(* IEC 61131-3 sources: JingjiangArm/moonboxpro_arm_8.4/Application/Application/任务列表/LogTask/文件存储/数据存储&日志操作, 8 files *)

(* ---- ENUMS_TIMEFORMAT.st ---- *)
(*@CES
Name=ENUMS_TIMEFORMAT
Type=Gvl
TypeGuid=2db5746d-d284-4425-9f7f-2663a34b0ebc
Guid=3fd86c5d-f4c2-4e63-8cc9-6ae2cca08ccd
HasDeclaration=True
HasImplementation=False
*)
{DECLARATION}
//{attribute 'qualified_only'}
//{attribute 'strict'}
TYPE ENUMS_TIMEFORMAT : (
	TIMEFORMAT_NO_HYPHEN		, (* yyyymmddHHMMSS *)
	TIMEFORMAT_HYPHEN_COLON		, (* yyyy-mm-dd HH:MM:SS *)
	TIMEFORMAT_HYPHEN_DOT		, (* yyyy.mm.dd.HHMMSS *)
	TIMEFORMAT_MMDD				, (* mmdd *)
	TIMEFORMAT_MMDDHH			  (* mmddHH *)
);
END_TYPE
{IMPLEMENTATION}

(* ---- StAxisWatchDetails.st ---- *)
(*@CES
Name=StAxisWatchDetails
Type=Gvl
TypeGuid=2db5746d-d284-4425-9f7f-2663a34b0ebc
Guid=06521707-3ba7-4049-9244-d2161cd79c22
HasDeclaration=True
HasImplementation=False
*)
{DECLARATION}
{attribute 'pack_mode' := '1'}
TYPE StAxisWatchDetails :
STRUCT
// 	iStationId						: INT;(*主控站ID*)
// 	rGirth 							:REAL ; (*周长*)
// 	iRtn_Station					: INT;//返回值
// 	iRunMode_Station				: INT;//运动模式-3电子齿轮4龙门
// 	rPos_Prf						: REAL;//规划位置
// 	rPos_Enc						: REAL;//编码器位置
// 	rVel_Enc						: REAL;//编码器速度
// 	rTorque							: REAL;//扭矩输出
// 	rGantry_Err						: REAL;//龙门错误吗
//  	rTemperaTure					: REAL;//电机温度
// 	dwErr_Driver					: DWORD;//驱动器报警状态
// 	wSts_Driver						: WORD;//驱动器状态
// 	wSts_NetPort					: WORD;//端口状态
// 	wSts_NetRun						: WORD;//端口运行状态
//  	iErr_NetPort_a					: INT;//A误码率
//  	iErr_NetPort_b					: INT;//B误码率
// 	dwMotion_Sts					: DWORD;//运型状态
// 	uiVirtual_Cnt					: UINT;//虚拟码盘基数
// 	wVirtual_Sts					: WORD;//虚拟马盘状态
// 	uiBrake_Cnt						: UINT;//制动次数
// 	rCurrent_Driver					: REAL;//电流
// 	rVdc							: REAL;//母线电压
// 	uiStationType					: UINT;//站类型
// 	uiDrvParam_Imax					: UINT;(* 驱动参数|最大电流 *)
// 	uiDrvParam_Nrs					: UINT;(* 驱动参数|额定转速 *)
// 	uiDrvParam_Nos					: UINT;(* 驱动参数|过速转速 *)
// 	iDrvParam_PosOfst				: INT;(* 驱动参数|位置偏移 *)

	rGirth: REAL; (* 轴周长 *)
	lrPT_Pos: LREAL; (* 轴PT规划P *)
	diPT_Time: DINT; (* 轴PT规划T *)
	byPT_Type: BYTE; (* 轴PT段选择|2.PT_SEGMENT_NORMAL;1.PT_SEGMENT_EVEN;0.others *)
	rtnSts: INT; (* 返回状态 *)
	bySpace: BYTE; (* fifo空间 *)
	pfr: DWORD; (* 规划位置 *)
	enc_Lo16: INT; (* StPTSts.enc的低16位_跟随误差的低16位 *)
	driverSts: INT; (* 驱动器状态 *)
	driverErr: INT; (* 驱动器错误 *)
	netPortErr_a: INT; (* A口误码率 *)
	netPortErr_b: INT; (* B口误码率 *)
	motionSts: DWORD; (* 运动器状态 *)
	modal: WORD; (* 模态 *)
	brakeCnt: WORD; (* 制动电阻次数 *)
	driverCurrent: WORD; (* 驱动器电流 *)
	rVel_Axis: REAL; (* 轴速度 *)
	rAI_Axis_Coating: REAL; (* 当前值-中位值 *)
	enc_Hi16: WORD; (* StPTSts.enc的高16位_网络锁存时间的低16位 *)(* 新增14个字节|@2020.10.13.171810_ *)
	temperature: INT; (* 电机温度 *)
	vel: INT; (* 规划速度 *)
	netPortSts: INT; (* 网络端口连接状态 *)
	netRunSts: INT; (* 网络运行状态 *)
	virtualCnt: WORD; (* 虚拟码盘计数 *)
	virtualSts: WORD; (* 虚拟码盘状态 *)
	(*2022.5.25.131916 增加了锁存编码器值的保存*)
	dwCurAxisEnc_Lock: DWORD;(*当前轴锁存编码器值*)
	dwCurAxisSystime_Lock					: DWORD;(*当前轴锁存系统时间*)
(*2022.6.24.151851  取消使用*)
(*
	dwLastLinkageAxisEnc_Lock				: DWORD;(*上个联动轴锁存编码器值*)
	dwLastLinkageAxisSystime_Lock			: DWORD;(*上个联动轴锁存系统时间*)
*)
	(*2022.6.24.151255*)
	iai1_New16D:			INT;(*模拟量输入1*)
	iai2_New16D:			INT;(*温控输入*)
	rDc_Voltage:REAL;(*母线电压值*)
	idriverErr_H: INT; (* 驱动器错误 |高16bit*)

	(*新增加的单联动切换功能，在出现问题的时候为了方便查找问题,增加了文件保存内容*)
	(*电机使能模式|0: 不使能 1: 使能 3: 使能后轴可以手动转动 4: 取消模式3状态
	3、4以为的值都不允许set
	实际应用下会3、4状态下切换*)
	wEnableMode_Motor						: WORD;
	byEnableModeSwitchDne					: BYTE;(*使能模式切换成功了|.0 =3 成功了
																		.1 =4 成功了*)
	xMoveEnable_Motor						: BOOL;(*电机运动使能|用于控制驱动器是否进行电机控制|与单联动比较切换电机是否运动*)

	byAxisMotionSts:BYTE;(*轴运动状态标志|0:同步运动状态.
										  |1:同步运动时停止运动状态.
										  |2:停止运动状态
										  |3:停止运动时加速到单运行速度状态.
										  |4:单运行时减速到停止状态.
										  |5:停止运动时或者使用单运行速度运行时加速到同步运动状态.
										  |6:非同步运动时急停到0状态.
										  |7:非同步运动时空转停机到0状态.*)
(*2022.10.22.162829保存加热相关数据*)
	rPIDValue:REAL;(*pid计算调整量*)
	rPV_Unit:REAL;(*当前温度*)
	rSV_Unit:REAL;(*设定温度*)
	rValue_P:REAL;
	rValue_I:REAL;
	rValue_D:REAL;
	iNumCount:INT;

(*end_2022.10.22.163310*)

END_STRUCT
END_TYPE

{IMPLEMENTATION}

(* ---- StRecord_A.st ---- *)
(*@CES
Name=StRecord_A
Type=Gvl
TypeGuid=2db5746d-d284-4425-9f7f-2663a34b0ebc
Guid=136b24a0-c4f1-416e-bf48-48716262a31a
HasDeclaration=True
HasImplementation=False
*)
{DECLARATION}
{attribute 'pack_mode' := '1'}
TYPE StRecord_A :
STRUCT
	dwCurYMD: DWORD;
	dwCurHMSU: DWORD;
	byAxisId: BYTE; (* 轴id *)
	byGrpId: BYTE; (* 系id *)
	uiNum: UINT; (* 减速比分子 *)
	uiDen: UINT; (* 减速比分母 *)
	udiVel: UDINT; (* 主机速度|单位:0.01m/min *)
	udiGirth: UDINT; (* 版周长|单位:0.001mm *)
	iGateSa: INT; (* 波门地址1 *)
	iGateSaEx: INT; (* 波门地址2 *)
	byMarkTypeId: BYTE; (* 标记形式 *)
	byMarkArrangeId: BYTE; (* 标记排列 *)
	wSwitchRef: WORD; (* 开关状态 *)
	wStatusRef: WORD; (* 手/自动状态 *)
	wExtendedProf: WORD;
			(* 描述位|
				bit0=1表示合压中,
				bit1=1标识等料长,
				bit2=1标识裁切让料头

				bit8=1表示第一组波门T1极性
				bit9=1表示第一组波门T2极性
				bit10=1表示第二组波门T1极性
				bit11=1表示第二组波门T2极性
*)
	byStsV: BYTE; (* 纵向误差状态 *)
	byStsH: BYTE; (* 横向误差状态 *)
	aiKpid_setup_v: ARRAY [1..3] OF INT; (*界面设置的纵向pid*)
	aiKpid_setup_h: ARRAY [1..3] OF INT; (*界面设置的横向pid*)
	aiKpid_used_v: ARRAY [1..3] OF INT; (*使用中的纵向pid*)
	aiAdjVal_vh: ARRAY [1..2] OF INT; (*纵横向版修正量*)
	lrFilmLengthFromPrevUnit: LREAL; (* 预套准料长总值 *)
	byCouplingMask: BYTE; (* 耦合开关 *)
	iErrDataRelay_Index_V: INT; (* 取的误差间隔幅数 *)
	iErrDataRelay_V: INT; (* 传来的误差 *)
	aiErrorVal_vh: ARRAY [1..2] OF INT; (*纵横向误差*)
	aiAdjValCalcByPid_vh: ARRAY [1..2] OF INT; (*计算的调整量*)

	alrCurCycleAdjustVal_Auto_vh: ARRAY [1..2] OF LREAL; (* 自动调整*)
	alrCurCycleAdjustVal_Rapid_vh: ARRAY [1..2] OF LREAL; (* 快速对版调整*)
	alrCurCycleAdjustVal_ManuCoarse_vh: ARRAY [1..2] OF LREAL; (* 手动粗调*)
	alrCurCycleAdjustVal_ManuFine_vh: ARRAY [1..2] OF LREAL; (* 手动细调*)
	alrCurCycleAdjustVal_Coupling_vh: ARRAY [1..2] OF LREAL; (* 耦合量*)
	alrCurcycleAdjustVal_Compensate_vh: ARRAY [1..2] OF LREAL; (* 补偿量*)

	alrTotalAdjustVal_Auto_vh: ARRAY [1..2] OF LREAL; (* 自动调整仓库*)
	alrTotalAdjustVal_Rapid_vh: ARRAY [1..2] OF LREAL; (* 快速对版仓库*)
	alrTotalAdjustVal_ManuCoarse_vh: ARRAY [1..2] OF LREAL; (* 手动粗调仓库*)
	alrTotalAdjustVal_ManuFine_vh: ARRAY [1..2] OF LREAL; (* 手动细调仓库*)
	alrTotalAdjustVal_Coupling_vh: ARRAY [1..2] OF LREAL; (* 耦合量仓库*)
	alrTotalAdjustVal_Compensate_vh: ARRAY [1..2] OF LREAL; (* 补偿量仓库*)

	alrExecutedAdjVal_Auto_vh: ARRAY [1..2] OF LREAL; (* 已经执行的自动调整量*)
	alrExecutedAdjVal_Rapid_vh: ARRAY [1..2] OF LREAL; (* 已经执行的快速调整量*)
	alrExecutedAdjVal_ManuCoarse_vh: ARRAY [1..2] OF LREAL; (* 已经执行的手动粗调量*)
	alrExecutedAdjVal_ManuFine_vh: ARRAY [1..2] OF LREAL; (* 已经执行的手动细调量*)
	alrExecutedAdjVal_Coupling_vh: ARRAY [1..2] OF LREAL; (* 已经执行的耦合量*)
	alrExecutedAdjVal_Compensate_vh: ARRAY [1..2] OF LREAL; (* 已经执行的补偿量*)

	dwFS_index: DWORD; (* 精采样数据幅数索引 *)
	aiParsing_base: ARRAY [1..2] OF INT; (* 两路信号基线 *)
	aiParsing_min: ARRAY [1..2] OF INT; (* 两路信号最小值 *)
	aiParsing_max: ARRAY [1..2] OF INT; (* 两路信号最大值 *)
	dwIndex:DWORD; (* 索引号，用于与张力数据对应*)
	(*保存精采样标志@可能会滞后一幅*)
	xSaveFineSampleData_ToArc:BOOL;

	(*2023.09.04.092458  增加*)
	aiActErrorVal_vh: ARRAY [1..2] OF INT; (*纵横向误差原始值|未经过平均的*)

	(*计算的当前误差@8bytes*)
	iVerror_FollowPreUnit 					: INT; (*纵向跟前一色误差@05号命令*)
	iVerror_Follow1Unit 					: INT;(*纵向跟1色误差@05号命令*)
	iHerror_FollowPreUnit 					: INT; (*横向跟前一色误差@05号命令*)
	iHerror_Follow1Unit 					: INT;(*横向跟1色误差@05号命令*)

	(*2024.03.10.233250 修改*)
	rFinalAdjust_V_Act:REAL;(*小黄耦合函数输出的实际调整量@上一拍的值|2023.11.18.194816*)
	(*2026.5.7.175735套色算法测试lhy+*)
	dwTime:DWORD; (*2026.1.17.112058*)
	abyReserved:ARRAY [1..2] OF BYTE;
	(*2023.11.18.194736|+rFinalAdjust_V_Act@10-->6*)
(*2023.11.18.194636 屏蔽使用@使用上面的数组保持内存对其|保证解析工具的兼容*)
(*
	(*2023.09.11.104053 增加误差滤波函数的数据保存*)
	iCurrentObservationError : INT;(*当前观测误差*)
	iPreviousAdjustment : INT;(*上一幅调整量@正误差需要输入负调整量-外面根据正逆序修改*)
	(*最终返回预测误差*)
	iPredictionError : INT; (*预测误差*)
	rKalmanGain:REAL;(*增益*)
*)

END_STRUCT
END_TYPE

{IMPLEMENTATION}

(* ---- StRecord_T.st ---- *)
(*@CES
Name=StRecord_T
Type=Gvl
TypeGuid=2db5746d-d284-4425-9f7f-2663a34b0ebc
Guid=143e99cc-3331-46fe-a10c-279acbbec24f
HasDeclaration=True
HasImplementation=False
*)
{DECLARATION}
{attribute 'pack_mode' := '1'}
TYPE StRecord_T :
STRUCT
	dwYMD: DWORD;(* 年月日*)
	dwHMSU: DWORD;(* 时分秒毫秒*)
	byGrpId: BYTE; (* 系id\自动赋值 *)
	dwIndex: DWORD; (* 主任务周期索引 *)
	rVel_Cur: REAL; (* 当前速度 *)
	rVel_Film: REAL; (* 料膜速度 *)
	uiMillimeter_Diam_PaperTube_Uw: UINT; (* 放料卷纸卷直径|单位mm|2019.11.28.112452 *)
	uiMicron_FilmThickness: UINT; (* 料膜厚度|单位um|2019.11.28.112452 *)
	uiMicron_FilmThickness_RevCalculated: UINT; (* 料膜厚度的反算值|单位um|2019.11.29.153103 *)
	uiMeterLength_SurplusMaterial: UINT; (* 剩余料膜长度|单位m|2019.11.28.112452 *)
	dwFlag: DWORD; (* 标志位*)
					(*bit.0:放料当前轴
					  bit.1:收料当前轴
					  bit.2:压力传感器使能
					  bit.16:放料翻转架正转
					  bit.17:放料翻转架反转
					  bit.18:收料翻转架正转
					  bit.19:收料翻转架反转
					  bit.20:放料A轴正转使能
					  bit.21:放料B轴正转使能
					  bit.22:收料A轴正转使能
					  bit.23:收料B轴正转使能
					  bit.26:放料预估弧面信号
					  bit.27:放料对射电眼信号输入
					  bit.28:放料裁切按钮输入
					  bit.29:放料弧面信号输入
					  bit.30:放料裁刀输出
					  bit.31:放料胶辊输出
					*)
	arAI_UwRw_IfOf: ARRAY [1..4] OF REAL; (* 摆臂输入|rAI_Uw|rAI_Rw|rAI_If|rAI_Of *)
	arPI_UwRw_IfOf: ARRAY [1..4] OF REAL; (* Pi计算量|rPi_Uw|rPi_Rw|rPi_If|rPi_Of *)
	arDiam_UwRw_Girth_IfOf: ARRAY [1..4] OF REAL; (* 周长或直径|rGirth_Uw|rGirth_Rw|rGirth_If|rGirth_Of *)
	arStep_UwRw_IfOf: ARRAY [1..4] OF REAL; (* 前馈|rStep_Uw|rStep_Rw|rStep_If|rStep_Of *)
	arVel_UwRw_IfOf: ARRAY [1..4] OF REAL; (* 速度|rVel_Uw|rVel_Rw|rVel_If|rVel_Of *)
(*收放料PID保存改为*100||保留精度-改word型*)
	aiKpid_UwRw_IfOf: ARRAY [1..4,1..3] OF WORD; (* Kpid参数|iP_Uw|iI_Uw|iD_Uw|......|iP_Of|iI_Of|iD_Of *)
	rPressure_Tar: REAL; (* 压力传感器目标压力*)
	rCurPressureValue: REAL; (* 压力传感器实时压力*)
	wAOVolt_If_inverter: WORD; (* 放牵模拟量输出*)
	wAOVolt_Of_inverter: WORD; (* 收牵模拟量输出*)
	rStdVol_AI_cur: REAL; (* 当前卷径电压 *)
	rStdVol_AI_use: REAL; (* 计算用的卷径电压 *)
	rDia_New_Auto: REAL; (* 计算所得新卷卷径*)
	rUwPreVel_Vol_A: REAL; (* 放料预驱速度电压*)
	rUwPreVel_Vol_B: REAL; (* 放料预驱速度电压*)
	rRwPreVel_Vol_A: REAL; (* 收料预驱速度电压*)
	rRwPreVel_Vol_B: REAL; (* 收料预驱速度电压*)
	rUwPreVel: REAL; (* 放料预驱速度*)
	rRwPreVel: REAL; (* 收料预驱速度*)
	iMotionStepId: INT; (* MOTION_STEP_... *)
	iPromptMsgId: INT; (* 报警代码*)
	wPreHotRollerFrq: WORD; (* 预热辊输出*)
	wWaterCoolRollerFrq: WORD; (* 水冷辊输出*)
	byPlcLoad: BYTE; (* cpu消耗|2020.4.14.153153 *)
(*2023.09.20.134044 为了保证兼容|将这两个不用的real型变量作为他用|保证解析工具的内存对其*)
(*
	rVel_SelfAdjust_Uw_A: REAL; (* 2020.10.8.164751|放料A轴自调整速度 *)
	rVel_SelfAdjust_Uw_B: REAL; (* 2020.10.8.164751|放料B轴自调整速度 *)
*)
	awPressRollerVol:ARRAY [1..4] OF WORD;(*压力传感器电压值@留出来4个*)

	(*2021.8.27.170829 增加放料翻转架需要保存的变量*)
	rTowerThetaCur_Uw:REAL;
	rDeltaW_RPMIN_Uw:REAL;
	rFilmToTowerRollerDis: REAL;(*料膜距离导向辊距离|mm*)

	(*2021.8.27.093201  卷径估计需要变量保持*)
	rEstiDia_Uw:REAL;(*放料卷径估计值*)
	rEstiThickNess_Uw:REAL;(*放料厚度估计值*)
	rMainVel_Uw:REAL;(*卷径估计使用时 放料主速度*)
	rEstiDia_Rw:REAL;(*收料卷径估计值*)
	rEstiThickNess_Rw:REAL;(*收料厚度估计值*)
	rMainVel_Rw:REAL;(*卷径估计使用时 收料主速度*)

	(*2021.9.13.161022*)
(*2024.7.12.113636 复用位置*)
(*
	(*放料接料补偿-窄方波+微分*)
	rSpliceCompensate_Uw:REAL;(*计算的补偿值*)
	rSpliceCompensate_Wr_Uw:REAL;(*裁切补偿实际写入的值*)
*)
	rUseDiamWuCompensate_Uw:REAL;(*放料张力算法计算使用的卷径值*)
	rUseDiamWuCompensate_Rw:REAL;(*收料张力算法计算使用的卷径值*)

	(*2022.9.7.215546增加了锥度值的数据存储|单位0.01*)
	uiTaper_Cur_Uw:UINT;
	uiTaper_Cur_Rw:UINT;
	uiTaper_Cur_If:UINT;
	uiTaper_Cur_Of:UINT;

(*2022.10.22.162829保存加热相关数据*)
	iPidAlgorithm_Threshold:INT;(*温控PDI介入阀值*)
	iMaxOutValue:INT;(*温控最大调整量*)
	rKp:REAL;
	rKi:REAL;
	rKd:REAL;
	uiCtlCycle_Ms:UINT;(*调整周期*)
(*end2022.10.22.163043*)

	(*2022.11.2.104744 增加了伪随机测试需要的*)
	byRoundTime:BYTE;
	rVolAdditionValue:REAL;(*随机数的值*)
	rAmplitude:REAL;(*伪随机幅值*)

	(*2023.09.18.182952 同步*)
	(*2023.09.08.155701 增加*)
	rWuCompensate_Uw:REAL;(*补偿的转速(R/MIN)|计算的*)
	rDh_Uw:REAL;(*扰动的估计值(M/S)|计算的*)
	rWuCompensate_Act_Uw:REAL;(*补偿的转速(R/MIN)|实际使用的*)

	(*2024.7.11.134605+*)
	rEstiDia_LowPass_Uw:REAL;(*放料低通后卷径值*)
	byKalmanFilterType_Rw:BYTE;(*收料卡尔曼估计的方式值*)
	rWc_LowPass_Diam_Rw:REAL;(*收料卷径截止频率值*)
	rWuCompensate_Rw:REAL;(*补偿的转速(R/MIN)|计算的*)
	rWuCompensate_Act_Rw:REAL;(*补偿的转速(R/MIN)|实际使用的*)
	rKc_Rw:REAL;(*收料补偿值增益|卡尔曼估计方式1 2 3 4 5*)
	rEstiDia_LowPass_Rw:REAL;(*收料低通后卷径值*)
	(*2024.9.10.122313+8bytes*)
	rAntiNotch_Out_If:REAL;(*放牵摆臂过陷波值*)
	rAntiNotch_Out_Uw:REAL;(*放料摆臂过陷波值*)
	abyReserved_11:ARRAY [1..3] OF BYTE;(*2024.7.3.153430 替换了|将来作为别的用途*)
					(*rAntiNotch_Out_If-->rAntiNotch_Out_Uw|11->3*)
					(*rEstiDia_LowPass_Uw-->rEstiDia_LowPass_Rw|36->11*)

	xSaveFineSampleData:BOOL;(*2023.5.29.105143@精采样存储按钮|2023.6.13.090435*)

	(*2024.01.11.153854 增加了一些张力控制器的参数保存*)
	rWc_LowPass_Diam_Uw:REAL;(*放疗卷径截止频率值*)
	byKalmanFilterType_Uw:BYTE;(*放料卡尔曼估计的方式值*)
	rKc_Uw:REAL;(*放料补偿值增益|卡尔曼估计方式1 2 3 4 5*)
(*	rKc_1_Uw:REAL;(*放料补偿值增益|卡尔曼估计方式0*)*)
	abySpace_0:ARRAY [1..4] OF BYTE;(*增加空余部分*)

	(*2024.01.11.153922 任务执行周期数据保存*)
	byCycleTime_PlcPrg		: BYTE;(* 任务消耗时间 *)
	byIntervalTime_PlcPrg	: BYTE;(* 任务间隔 *)

(*	bya_Youla_Uw:BYTE;(*youla控制器的系统参数a@保留0.1|支持最大值25.5*)*)

	abySpace_1:ARRAY [1..1] OF BYTE;(*增加空余部分*)

	byTotalVariableAxisNum: BYTE; (* 轴数量 *)
	dwMask_VariableAxisDetails: DWORD; (* bit0=Axis.1|bit31=Axis.32 *)
END_STRUCT
END_TYPE
{IMPLEMENTATION}

(* ---- StTravelDataItem.st ---- *)
(*@CES
Name=StTravelDataItem
Type=Gvl
TypeGuid=2db5746d-d284-4425-9f7f-2663a34b0ebc
Guid=62504b07-d26b-473c-be85-27d686726a0a
HasDeclaration=True
HasImplementation=False
*)
{DECLARATION}
TYPE StTravelDataItem :
STRUCT
	uiValidBytesNum		: UINT;(* 描述abyPayload有效的字节数量 *)
	abyPayload			: ARRAY [1..BYTES_PER_ROW_RECORD] OF BYTE;
END_STRUCT
END_TYPE

{IMPLEMENTATION}

(* ---- StTravelDataRec.st ---- *)
(*@CES
Name=StTravelDataRec
Type=Gvl
TypeGuid=2db5746d-d284-4425-9f7f-2663a34b0ebc
Guid=4a1c87c8-507f-49a1-a6b5-dfc3139d89be
HasDeclaration=True
HasImplementation=False
*)
{DECLARATION}
TYPE StTravelDataRec :
STRUCT
	uiWR				: UINT;(* 写位置 *)
	uiRD				: UINT;(* 读位置 *)
	astStTravelDataItem	: ARRAY [1..MAX_ROWS_OF_RECORD] OF StTravelDataItem;(* 数据静荷区域 *)
END_STRUCT
END_TYPE
{IMPLEMENTATION}

(* ---- StTravelLogItem.st ---- *)
(*@CES
Name=StTravelLogItem
Type=Gvl
TypeGuid=2db5746d-d284-4425-9f7f-2663a34b0ebc
Guid=d92a6104-9117-400f-b58f-f96bab8fae06
HasDeclaration=True
HasImplementation=False
*)
{DECLARATION}
TYPE StTravelLogItem :
STRUCT
	wLogLevelId				: WORD;(* 参考LOG_LEVEL_xxx *)
	sInfo					: STRING(256);
END_STRUCT
END_TYPE

{IMPLEMENTATION}

(* ---- StTravelLogRec.st ---- *)
(*@CES
Name=StTravelLogRec
Type=Gvl
TypeGuid=2db5746d-d284-4425-9f7f-2663a34b0ebc
Guid=1e9822ea-ea5b-4373-ab67-94f283ee71ec
HasDeclaration=True
HasImplementation=False
*)
{DECLARATION}
TYPE StTravelLogRec :
STRUCT
	uiIndex_Wr: UINT;(* 当前写入位置 *)
(*	uiIndex_Peek: UINT;(* 当前窥探位置 *)*)
	uiIndex_Rd: UINT;(* 当前读取位置 *)
	xOverwrite: BOOL;(* 过圈标志 *)
	astStTravelLogItem: ARRAY [1..GC_LOG_ITEM_MAX_NUM] OF StTravelLogItem;(* 日志队列 *)
END_STRUCT
END_TYPE
{IMPLEMENTATION}
